Fanuc KAREL source: KT00736.KL

PROGRAM KT00736
%NOLOCKGROUP
VAR
  ARG: ARRAY[4] OF STRING[20]
  OUT: BOOLEAN
BEGIN
  OUT = UNINIT(ARG)
END KT00736
